	110: //Verifica se a reta indexada é a última criada
		IF NOT IHM.CutMode THEN
			IF PLC.CutLine = PLC.Grid THEN
				Auto.State := 118;
				ELSIF PLC.CutLine <> PLC.Grid THEN
					Auto.State := 111;
			END_IF
			ELSIF IHM.CutMode THEN
				IF PLC.CutLine = PLC.GridDesigner_LastLine THEN
					Auto.State := 118;
					ELSIF PLC.CutLine <> PLC.GridDesigner_LastLine THEN
						Auto.State := 111;
				END_IF
		END_IF
	
	111: //Passa para próxima reta
		PLC.CutLine := PLC.CutLine + 1;
		Auto.State := 30;
	
	118: //Recebe valor da última reta do eixo da altura ou primeira reta do eixo da largura
		IF NOT IHM.CutMode THEN
			PLC.CutLine := PLC.GridDesigner_LastLine;
			Auto.State := 119;
			ELSIF IHM.CutMode THEN
				PLC.CutLine := 21;
				Auto.State := 119;
		END_IF
	
	119: //Serra 90° ou 0° + Serra Ligada
		IF NOT IHM.CutMode THEN
			PLC.Axis[4].OperationDistance := 0;
			Auto.State := 120;
			ELSIF IHM.CutMode THEN
				PLC.Axis[4].OperationDistance := 90;
				Auto.State := 120;
		END_IF
	
	120: //Movimenta eixo W
		PLC.Axis[4].OperationStart := TRUE;
		IF NOT PLC.Axis[4].OperationDone THEN
			Auto.State := 121;
		END_IF
	
	121: //Aguarda movimentação do eixo
		IF PLC.Axis[4].OperationDone THEN
			PLC.Axis[4].OperationStart := FALSE;
			Auto.State := 122;
		END_IF
	
	122: //Posicão Zero Peça X (descontando borda de entrada) + Zero Peça Y da peça indexada
		IF NOT IHM.CutMode THEN
			PLC.Axis[1].OperationDistance := PLC.OrthogonalPieces[PLC.CutLine].LastVertexAbsX + (IHM.PrEntryEdgeX * -1);
			PLC.Axis[2].OperationDistance := PLC.OrthogonalPieces[PLC.CutLine].ZeroPieceY;
			PLC.Axis[1].OperationAbsolute := TRUE;
			PLC.Axis[2].OperationAbsolute := TRUE;
			Auto.State := 130;
			ELSIF IHM.CutMode THEN
				PLC.Axis[1].OperationDistance := PLC.OrthogonalPieces[PLC.CutLine].ZeroPieceX;
				PLC.Axis[2].OperationDistance := PLC.OrthogonalPieces[PLC.CutLine].ZeroPieceY + IHM.PrEntryEdgeY;
				PLC.Axis[1].OperationAbsolute := TRUE;
				PLC.Axis[2].OperationAbsolute := TRUE;
				Auto.State := 130;
		END_IF
	
	130: //Movimenta eixo X
		PLC.Axis[1].OperationStart := TRUE;
		IF NOT PLC.Axis[1].OperationDone THEN
			Auto.State := 131;
		END_IF
	
	131: //Movimenta eixo Y
		PLC.Axis[2].OperationStart := TRUE;
		IF NOT PLC.Axis[2].OperationDone THEN
			Auto.State := 132;
		END_IF
	
	132: //Aguarda movimento 90°/0° e movimentações de X e Y
		IF NOT IHM.CutMode AND PLC.Axis[4].Position = 0 OR IHM.CutMode AND PLC.Axis[4].Position = 90 THEN
			IF PLC.Axis[1].OperationDone AND PLC.Axis[2].OperationDone THEN
				PLC.Axis[1].OperationStart := FALSE;
				PLC.Axis[2].OperationStart := FALSE;
				Auto.State := 140;
			END_IF
		END_IF
	
	140: //Posição dentro da peça
		PLC.Axis[3].OperationDistance := IHM.PrInsidePiece;
		PLC.Axis[3].OperationAbsolute := TRUE;
		Auto.State := 150;
	
	150: //Movimenta eixo Z
		PLC.Axis[3].OperationStart := TRUE;
		IF NOT PLC.Axis[3].OperationDone THEN
			Auto.State := 151;
		END_IF
	
	151: //Aguarda movimentação do eixo
		IF PLC.Axis[3].OperationDone THEN
			PLC.Axis[3].OperationStart := FALSE;
			Auto.State := 160;
		END_IF
	
	160: //Deslocamento da largura (descontando bordas de entrada e saída) da peça indexada
		IF NOT IHM.CutMode THEN
			PLC.Axis[1].OperationDistance := (PLC.OrthogonalPieces[PLC.CutLine].Lenght * -1) + IHM.PrEntryEdgeX + IHM.PrLeadingEdgeX;
			PLC.Axis[1].OperationAbsolute := FALSE;
			Auto.State := 170;
			ELSIF IHM.CutMode THEN
				PLC.Axis[2].OperationDistance := PLC.OrthogonalPieces[PLC.CutLine].Lenght + (IHM.PrEntryEdgeY * -1) + (IHM.PrLeadingEdgeY * -1);
				PLC.Axis[2].OperationAbsolute := FALSE;
				Auto.State := 170;
		END_IF
	
	170: //Movimenta X ou Y
		IF NOT IHM.CutMode THEN
			PLC.Axis[1].OperationStart := TRUE;
			IF NOT PLC.Axis[1].OperationDone THEN
				Auto.State := 171;
			END_IF
			ELSIF IHM.CutMode THEN
				PLC.Axis[2].OperationStart := TRUE;
				IF NOT PLC.Axis[2].OperationDone THEN
					Auto.State := 171;
				END_IF
		END_IF
	
	171: //Aguarda movimentação X ou Y
		IF NOT IHM.CutMode AND PLC.Axis[1].OperationDone THEN
			PLC.Axis[1].OperationStart := FALSE;
			Auto.State := 180;
			ELSIF IHM.CutMode AND PLC.Axis[2].OperationDone THEN
				PLC.Axis[2].OperationStart := FALSE;
				Auto.State := 180;
		END_IF
	
	180: //Posição fora da peça
		PLC.Axis[3].OperationDistance := IHM.PrOutsidePiece;
		PLC.Axis[3].OperationAbsolute := TRUE;
		Auto.State := 190;
	
	190: //Movimenta eixo Z
		PLC.Axis[3].OperationStart := TRUE;
		IF NOT PLC.Axis[3].OperationDone THEN
			Auto.State := 191;
		END_IF
	
	191: //Aguarda movimentação do eixo
		IF PLC.Axis[3].OperationDone THEN
			PLC.Axis[3].OperationStart := FALSE;
			Auto.State := 200;
		END_IF
	
	200: //Verifica se a reta indexada é a primeira
		IF NOT IHM.CutMode THEN
			IF PLC.CutLine = 0 THEN
				Auto.State := 1000;
				ELSIF PLC.CutLine <> 0 THEN
					Auto.State := 201;
			END_IF
			ELSIF IHM.CutMode THEN
				IF PLC.CutLine = PLC.Grid THEN
					Auto.State := 1000;
					ELSIF PLC.CutLine <> PLC.Grid THEN
						Auto.State := 202;
				END_IF
		END_IF
	
	201: //Passa para reta anterior
		PLC.CutLine := PLC.CutLine - 1;
		Auto.State := 122;
	
	202: //Passa para reta peça
		PLC.CutLine := PLC.CutLine + 1;
		Auto.State := 122;
	
	999: //Abortar rotina
		Automatic_Abort();
	
	1000: //Finalizar rotina
		Automatic_Done();
END_CASE
                    
END_ACTION

ACTION Cutting_Corner:
                      (*Condição para habilitar modo automático*)
IF PLC.Machine = States.Manual THEN
	IF IHM.btStart OR PLC.IO.Start THEN
		Auto.Start := TRUE;
		PLC.Machine := States.Automatic;
		Auto.State := 1;
	END_IF
	(*Condição para parar processo*)
	ELSIF PLC.Machine = States.Automatic THEN
		IF IHM.btStop OR PLC.IO.Stop OR PLC.Axis[1].Error OR PLC.Axis[2].Error OR PLC.Axis[3].Error OR PLC.Axis[4].Error THEN
			Auto.State := 999;
		END_IF
END_IF

(*Rotina de corte corner [L]*)
CASE Auto.State OF
	1: //Estado rodando
		Automatic_Running();
	
	2: //Reseta variaveis
		AutomaticCorner_Reverse := FALSE;
		PLC.CutStraight := 0;
		AutomaticCorner_CuttingStep := 0;
		Auto.State := 10;
	
	10: //Posição fora da peça
		PLC.Axis[3].OperationDistance := IHM.PrOutsidePiece;
		PLC.IO.SawSpin := TRUE;
		PLC.Axis[3].OperationAbsolute := TRUE;
		Auto.State := 11;
	
	11: //Movimenta eixo Z
		PLC.Axis[3].OperationStart := TRUE;
		IF NOT PLC.Axis[3].OperationDone THEN
			Auto.State := 12;
		END_IF
	
	12: //Aguarda movimntação do eixo
		IF PLC.Axis[3].OperationDone THEN
			PLC.Axis[3].OperationStart := FALSE;
			Auto.State := 20;
		END_IF
	
	20: //Serra 90°
		PLC.Axis[4].OperationDistance := 90;
		Auto.State := 21;
	
	21: //Movimenta eixo W
		PLC.Axis[4].OperationStart := TRUE;
		IF NOT PLC.Axis[4].OperationDone THEN
			Auto.State := 22;
		END_IF
	
	22: //Aguarda movimentação do eixo
		IF PLC.Axis[4].OperationDone THEN
			PLC.Axis[4].OperationStart := FALSE;
			Auto.State := 30;
		END_IF
	
	30: //Posicão Zero Peça X + Zero Peça Y (descontando borda de entrada) da peça indexada
		IF NOT AutomaticCorner_HorizontalCutting THEN
			PLC.Axis[1].OperationDistance := PLC.CornerPieces[PLC.CutStraight].ZeroPieceX;
			PLC.Axis[2].OperationDistance := PLC.CornerPieces[PLC.CutStraight].ZeroPieceY + PLC.CornerPieces[PLC.CutStraight].EntryEdge;
			PLC.Axis[1].OperationAbsolute := TRUE;
			PLC.Axis[2].OperationAbsolute := TRUE;
			Auto.State := 40;
			ELSIF AutomaticCorner_HorizontalCutting THEN
				PLC.Axis[1].OperationDistance := PLC.CornerPieces[PLC.CutStraight].LastVertexAbsX + (PLC.CornerPieces[PLC.CutStraight].EntryEdge * -1);
				PLC.Axis[2].OperationDistance := PLC.CornerPieces[PLC.CutStraight].ZeroPieceY;
				PLC.Axis[1].OperationAbsolute := TRUE;
				PLC.Axis[2].OperationAbsolute := TRUE;
				Auto.State := 40;
		END_IF
	
	40: //Movimenta eixo X
		PLC.Axis[1].OperationStart := TRUE;
		IF NOT PLC.Axis[1].OperationDone THEN
			Auto.State := 41;
		END_IF
	
	41: //Movimenta eixo Y
		PLC.Axis[2].OperationStart := TRUE;
		IF NOT PLC.Axis[2].OperationDone THEN
			Auto.State := 42;
		END_IF
	
	42: //Aguardaserra 90° ou 0° e movimentações do eixo X e Y
		IF (NOT AutomaticCorner_HorizontalCutting AND PLC.Axis[4].Position = 90 AND PLC.Axis[1].OperationDone AND PLC.Axis[2].OperationDone) OR (AutomaticCorner_HorizontalCutting AND PLC.Axis[4].Position = 90 AND PLC.Axis[1].OperationDone AND PLC.Axis[2].OperationDone) THEN
			PLC.Axis[1].OperationStart := FALSE;
			PLC.Axis[2].OperationStart := FALSE;
			Auto.State := 50;
		END_IF
	
	50: //Posição dentro da peça
		PLC.Axis[3].OperationDistance := IHM.PrInsidePiece;
		PLC.Axis[3].OperationAbsolute := TRUE;
		Auto.State := 60;
	
	60: //Movimenta eixo Z
		PLC.Axis[3].OperationStart := TRUE;
		IF NOT PLC.Axis[3].OperationDone THEN
			Auto.State := 61;
		END_IF
	
	61: //Aguarda movimentação do eixo
		IF PLC.Axis[3].OperationDone THEN
			PLC.Axis[3].OperationStart := FALSE;
			Auto.State := 70;
		END_IF
	
	70: //Deslocamento da altura (descontando bordas de entrada e saída) da peça indexada
		IF NOT AutomaticCorner_HorizontalCutting THEN
			PLC.Axis[2].OperationDistance := PLC.CornerPieces[PLC.CutStraight].Height + (PLC.CornerPieces[PLC.CutStraight].EntryEdge * -1) + (PLC.CornerPieces[PLC.CutStraight].LeadingEdge * -1);
			PLC.Axis[2].OperationAbsolute := FALSE;
			Auto.State := 80;
			ELSIF AutomaticCorner_HorizontalCutting THEN
				PLC.Axis[1].OperationDistance := (PLC.CornerPieces[PLC.CutStraight].Width * -1) + PLC.CornerPieces[PLC.CutStraight].EntryEdge + PLC.CornerPieces[PLC.CutStraight].LeadingEdge;
				PLC.Axis[1].OperationAbsolute := FALSE;
				Auto.State := 80;
		END_IF
	
	80: //Movimenta eixo X ou Y
		IF NOT AutomaticCorner_HorizontalCutting THEN
			PLC.Axis[2].OperationStart := TRUE;
			IF NOT PLC.Axis[2].OperationDone THEN
				Auto.State := 81;
			END_IF
			ELSIF AutomaticCorner_HorizontalCutting THEN
				PLC.Axis[1].OperationStart := TRUE;
				IF NOT PLC.Axis[1].OperationDone THEN
					Auto.State := 81;
				END_IF
		END_IF
	
	81: //Aguarda movimentação X ou Y
		IF NOT AutomaticCorner_HorizontalCutting AND PLC.Axis[2].OperationDone THEN
			PLC.Axis[2].OperationStart := FALSE;
			Auto.State := 90;
			ELSIF AutomaticCorner_HorizontalCutting AND PLC.Axis[1].OperationDone THEN
				PLC.Axis[1].OperationStart := FALSE;
				Auto.State := 90;
		END_IF
	
	90: //Posição fora de peça
		PLC.Axis[3].OperationDistance := IHM.PrOutsidePiece;
		PLC.Axis[3].OperationAbsolute := TRUE;
		Auto.State := 100;
	
	100: //Movimenta eixo Z
		PLC.Axis[3].OperationStart := TRUE;
		IF NOT PLC.Axis[3].OperationDone THEN
			Auto.State := 101;
		END_IF
	
	101: //Aguarda movimentação do eixo
		IF PLC.Axis[3].OperationDone THEN
			PLC.Axis[3].OperationStart := FALSE;
			Auto.State := 110;
		END_IF
	
	110: //Verifica espelhamento
		IF NOT IHM.CreationCorner_MirrorCorner THEN
			IF NOT AutomaticCorner_HorizontalCutting AND PLC.CutStraight = 2 THEN
				Auto.State := 111;
			END_IF
			IF (NOT AutomaticCorner_HorizontalCutting AND PLC.CutStraight <> 2) OR (AutomaticCorner_HorizontalCutting AND PLC.CutStraight <> 5) THEN
				Auto.State := 120;
			END_IF
			IF AutomaticCorner_HorizontalCutting AND PLC.CutStraight = 5 THEN
				Auto.State := 1000;
			END_IF
			ELSIF IHM.CreationCorner_MirrorCorner THEN
				IF NOT AutomaticCorner_HorizontalCutting AND PLC.CutStraight = 3 THEN
					Auto.State := 111;
				END_IF
				IF (NOT AutomaticCorner_HorizontalCutting AND PLC.CutStraight <> 3) OR (AutomaticCorner_HorizontalCutting AND PLC.CutStraight <> 8) THEN
					Auto.State := 120;
				END_IF
				IF AutomaticCorner_HorizontalCutting AND PLC.CutStraight = 8 THEN
					Auto.State := 1000;
				END_IF
		END_IF
	
	111: //Passa para próxima reta e gira serra para 0°
		AutomaticCorner_HorizontalCutting := TRUE;
		PLC.Axis[4].OperationDistance := 0;
		Auto.State := 112;
	
	112: //Movimenta eixo W
		PLC.Axis[4].OperationStart := TRUE;
		IF NOT PLC.Axis[4].OperationDone THEN
			Auto.State := 113;
		END_IF
	
	113: //Aguarda movimentação do eixo
		IF PLC.Axis[4].OperationDone THEN
			PLC.Axis[4].OperationStart := FALSE;
			Auto.State := 120;
		END_IF
	
	120: //Passa para próxima reta
		PLC.CutStraight := PLC.CutStraight + 1;
		Auto.State := 30;
	
	999: //Abortar rotina
		Automatic_Abort();
	
	1000: //Finaliza rotina
		Automatic_Done();
END_CASE
                    
END_ACTION

ACTION Cutting_Forms:
                      (*Condição para habilitar modo automático*)
IF PLC.Machine = States.Manual THEN
	IF IHM.btStart OR PLC.IO.Start THEN
		Auto.Start := TRUE;
		PLC.Machine := States.Automatic;
		Auto.State := 1;
	END_IF
	(*Condição para parar processo*)
	ELSIF PLC.Machine = States.Automatic THEN
		IF IHM.btStop OR PLC.IO.Stop OR PLC.Axis[1].Error OR PLC.Axis[2].Error OR PLC.Axis[3].Error OR PLC.Axis[4].Error THEN
			Auto.State := 999;
		END_IF
END_IF

(*Rotina de corte Formas*)
CASE Auto.State OF
	1: //Estado rodando
		Automatic_Running();
	
	2: //Reseta variaveis
		AutomaticForms_Segaments := 0;
		Auto.State := 10;
	
	10: //Posição fora da peça
		PLC.Axis[3].OperationDistance := IHM.PrOutsidePiece;
		PLC.Axis[3].OperationAbsolute := TRUE;
		PLC.IO.SawSpin := TRUE;
		Auto.State := 11;
	
	11: //Movimenta eixo Z
		PLC.Axis[3].OperationStart := TRUE;
		IF NOT PLC.Axis[3].OperationDone THEN
			Auto.State := 12;
		END_IF
	
	12: //Aguarda movimentação do eixo
		IF PLC.Axis[3].OperationDone THEN
			PLC.Axis[3].OperationStart := FALSE;
			Auto.State := 20;
		END_IF
	
	20: //Verifica qual figura foi selecionada
		IF IHM.Figure = 1 THEN
			Auto.State := 30; //Quadrado/Retangulo
			ELSIF IHM.Figure = 2 THEN
				Auto.State := 70; //Circulo
				ELSIF IHM.Figure = 3 THEN
					Auto.State := 50; //Hexagono
					ELSIF IHM.Figure = 4 THEN
						Auto.State := 60; //Triangulo
		END_IF

(*-----------------QUADRADO-----------------*)	
	
	30: //Gira serra 90°
		PLC.Axis[4].OperationDistance := 90;
		Auto.State := 31;
		
	31: //Movimenta eixo W
		PLC.Axis[4].OperationStart := TRUE;
		IF NOT PLC.Axis[4].OperationDone THEN
			Auto.State := 32;
		END_IF
	
	32: //Aguarda movimentação do eixo
		IF PLC.Axis[4].OperationDone THEN
			PLC.Axis[4].OperationStart := FALSE;
			Auto.State := 33;
		END_IF
	
	33: //Posição zero peça
		IF AutomaticForms_Segaments = 0 THEN
			PLC.Axis[1].OperationDistance := PLC.FormsSquare.ZeroPieceX;
			PLC.Axis[2].OperationDistance := PLC.FormsSquare.ZeroPieceY + IHM.PrEntryEdgeY;
			PLC.Axis[1].OperationAbsolute := TRUE;
			PLC.Axis[2].OperationAbsolute := TRUE;
			Auto.State := 34;
			ELSIF AutomaticForms_Segaments = 1 THEN
				PLC.Axis[1].OperationDistance := PLC.FormsSquare.LastVertexAbsX + IHM.SawThickness;
				PLC.Axis[2].OperationDistance := PLC.FormsSquare.ZeroPieceY + IHM.PrEntryEdgeY;
				PLC.Axis[1].OperationAbsolute := TRUE;
				PLC.Axis[2].OperationAbsolute := TRUE;
				Auto.State := 34;
		END_IF
	
	34: //Movimenta eixo X
		PLC.Axis[1].OperationStart := TRUE;
		IF NOT PLC.Axis[1].OperationDone THEN
			Auto.State := 35;
		END_IF
	
	35: //Movimenta eixo Y
		PLC.Axis[2].OperationStart := TRUE;
		IF NOT PLC.Axis[2].OperationDone THEN
			Auto.State := 36;
		END_IF
	
	36: //Aguarda movimento dos eixos e posição da serra 90°
		IF PLC.Axis[1].OperationDone AND PLC.Axis[2].OperationDone AND PLC.Axis[4].Position = 90 THEN
			PLC.Axis[1].OperationStart := FALSE;
			PLC.Axis[2].OperationStart := FALSE;
			Auto.State := 37;
		END_IF
	
	37: //Posição dentro da peça
		PLC.Axis[3].OperationDistance := IHM.PrInsidePiece;
		PLC.Axis[3].OperationAbsolute := TRUE;
		Auto.State := 38;
	
	38: //Movimenta eixo Z
		PLC.Axis[3].OperationStart := TRUE;
		IF NOT PLC.Axis[3].OperationDone THEN
			Auto.State := 39;
		END_IF
	
	39: //Aguarda movimentação do eixo
		IF PLC.Axis[3].OperationDone THEN
			PLC.Axis[3].OperationStart := FALSE;
			Auto.State := 40;
		END_IF
	
	40: //Deslocamento da altura
		PLC.Axis[2].OperationDistance := PLC.FormsSquare.Height + (IHM.PrEntryEdgeY * -1) + (IHM.PrLeadingEdgeY * -1);
		Auto.State := 41;
	
	41: //Movimenta eixo Y
		PLC.Axis[2].OperationStart := TRUE;
		IF NOT PLC.Axis[2].OperationDone THEN
			Auto.State := 42;
		END_IF
	
	42: //Aguarda movimento do eixo
		IF PLC.Axis[2].OperationDone THEN
			PLC.Axis[2].OperationStart := FALSE;
			Auto.State := 43;
		END_IF
	
	43: //Posição fora da peça
		PLC.Axis[3].OperationDistance := IHM.PrOutsidePiece;
		PLC.Axis[3].OperationAbsolute := TRUE;
		Auto.State := 44;
	
	44: //Movimento eixo Z
		PLC.Axis[3].OperationStart := TRUE;
		IF NOT PLC.Axis[3].OperationDone THEN
			Auto.State := 45;
		END_IF
	
	45: //Aguarda movimento do eixo
		IF PLC.Axis[3].OperationDone THEN
			PLC.Axis[3].OperationStart := FALSE;
			Auto.State := 46;
		END_IF
	
	46: //Soma na indexadora
		AutomaticForms_Segaments := AutomaticForms_Segaments + 1;
		Auto.State := 47;
	
	47: //Verifica se é o primeiro ou segundo corte
		IF AutomaticForms_Segaments = 2 THEN
			Auto.State := 48;
			ELSIF AutomaticForms_Segaments = 1 THEN
				Auto.State := 33;
		END_IF
	
	48: //Gira serra 0°
		PLC.Axis[4].OperationDistance := 0;
		Auto.State := 49;
		
	49: //Movimenta eixo W
		PLC.Axis[4].OperationStart := TRUE;
		IF NOT PLC.Axis[4].OperationDone THEN
			Auto.State := 50;
		END_IF
	
	50: //Aguarda movimentação do eixo
		IF PLC.Axis[4].OperationDone THEN
			PLC.Axis[4].OperationStart := FALSE;
			Auto.State := 51;
		END_IF
	
	51: //Posição zero peça
		IF AutomaticForms_Segaments = 2 THEN
			PLC.Axis[1].OperationDistance := PLC.FormsSquare.ZeroPieceX + IHM.PrEntryEdgeX;
			PLC.Axis[2].OperationDistance := PLC.FormsSquare.ZeroPieceY;
			Auto.State := 52;
			ELSIF AutomaticForms_Segaments = 3 THEN
				PLC.Axis[1].OperationDistance := PLC.FormsSquare.ZeroPieceX + IHM.PrEntryEdgeX;
				PLC.Axis[2].OperationDistance := PLC.FormsSquare.LastVertexAbsY + IHM.SawThickness;
				PLC.Axis[1].OperationAbsolute := TRUE;
				PLC.Axis[2].OperationAbsolute := TRUE;
				Auto.State := 52;
		END_IF
	
	52: //Movimenta eixo X
		PLC.Axis[1].OperationStart := TRUE;
		IF NOT PLC.Axis[1].OperationDone THEN
			Auto.State := 53;
		END_IF
	
	53: //Movimenta eixo Y
		PLC.Axis[2].OperationStart := TRUE;
		IF NOT PLC.Axis[2].OperationDone THEN
			Auto.State := 54;
		END_IF
	
	54: //Aguarda movimento dos eixos e posição da serra 0°
		IF PLC.Axis[1].OperationDone AND PLC.Axis[2].OperationDone AND PLC.Axis[4].Position = 0 THEN
			PLC.Axis[1].OperationStart := FALSE;
			PLC.Axis[2].OperationStart := FALSE;
			Auto.State := 55;
		END_IF
	
	55: //Posição dentro da peça
		PLC.Axis[3].OperationDistance := IHM.PrInsidePiece;
		PLC.Axis[3].OperationAbsolute := TRUE;
		Auto.State := 56;
	
	56: //Movimenta eixo Z
		PLC.Axis[3].OperationStart := TRUE;
		IF NOT PLC.Axis[3].OperationDone THEN
			Auto.State := 57;
		END_IF
	
	57: //Aguarda movimentação do eixo
		IF PLC.Axis[3].OperationDone THEN
			PLC.Axis[3].OperationStart := FALSE;
			Auto.State := 58;
		END_IF
	
	58: //Deslocamento da largura
		PLC.Axis[1].OperationDistance := PLC.FormsSquare.Width + (IHM.PrEntryEdgeX * -1) + (IHM.PrLeadingEdgeX * -1);
		Auto.State := 59;
	
	59: //Movimenta eixo Y
		PLC.Axis[1].OperationStart := TRUE;
		IF NOT PLC.Axis[1].OperationDone THEN
			Auto.State := 60;
		END_IF
	
	60: //Aguarda movimento do eixo
		IF PLC.Axis[1].OperationDone THEN
			PLC.Axis[1].OperationStart := FALSE;
			Auto.State := 61;
		END_IF
	
	61: //Posição fora da peça
		PLC.Axis[3].OperationDistance := IHM.PrOutsidePiece;
		PLC.Axis[3].OperationAbsolute := TRUE;
		Auto.State := 62;
	
	62: //Movimento eixo Z
		PLC.Axis[3].OperationStart := TRUE;
		IF NOT PLC.Axis[3].OperationDone THEN
			Auto.State := 63;
		END_IF
	
	63: //Aguarda movimento do eixo
		IF PLC.Axis[3].OperationDone THEN
			PLC.Axis[3].OperationStart := FALSE;
			Auto.State := 64;
		END_IF
	
	64: //Soma no indexador
		AutomaticForms_Segaments := AutomaticForms_Segaments + 1;
		Auto.State := 65;
	
	65: //Verifica se é o primeiro ou segundo corte
		IF AutomaticForms_Segaments = 4 THEN
			Auto.State := 1000;
			ELSIF AutomaticForms_Segaments = 3 THEN
				Auto.State := 51;
		END_IF
	
(*-----------------CIRCULO-----------------*)		
	
	70: //Gira serra 90°
		PLC.Axis[4].OperationDistance := 90;
		Auto.State := 71;
		
	71: //Movimenta eixo W
		PLC.Axis[4].OperationStart := TRUE;
		IF NOT PLC.Axis[4].OperationDone THEN
			Auto.State := 72;
		END_IF
	
	72: //Aguarda movimentação do eixo
		IF PLC.Axis[4].OperationDone THEN
			PLC.Axis[4].OperationStart := FALSE;
			Auto.State := 73;
		END_IF
	
	73: //Posição zero peça
		PLC.Axis[1].OperationDistance := PLC.FormsCircle.ZeroPieceX;
		PLC.Axis[2].OperationDistance := PLC.FormsCircle.Height / 2;
		PLC.Axis[1].OperationAbsolute := TRUE;
		PLC.Axis[2].OperationAbsolute := TRUE;
		Auto.State := 74;

	74: //Movimenta eixo X
		PLC.Axis[1].OperationStart := TRUE;
		IF NOT PLC.Axis[1].OperationDone THEN
			Auto.State := 75;
		END_IF
	
	75: //Movimenta eixo Y
		PLC.Axis[2].OperationStart := TRUE;
		IF NOT PLC.Axis[2].OperationDone THEN
			Auto.State := 76;
		END_IF
	
	76: //Aguarda movimento dos eixos e posição da serra 90°
		IF PLC.Axis[1].OperationDone AND PLC.Axis[2].OperationDone AND PLC.Axis[4].Position = 90 THEN
			PLC.Axis[1].OperationStart := FALSE;
			PLC.Axis[2].OperationStart := FALSE;
			Auto.State := 77;
		END_IF
	
	77: //Posição dentro da peça
		PLC.Axis[3].OperationDistance := IHM.PrInsidePiece;
		PLC.Axis[3].OperationAbsolute := TRUE;
		Auto.State := 78;
	
	78: //Movimenta eixo Z
		PLC.Axis[3].OperationStart := TRUE;
		IF NOT PLC.Axis[3].OperationDone THEN
			Auto.State := 79;
		END_IF
	
	79: //Aguarda movimentação do eixo
		IF PLC.Axis[3].OperationDone THEN
			PLC.Axis[3].OperationStart := FALSE;
			Auto.State := 80;
		END_IF
	
	80: //Primeira posição
		PLC.OperationAuxPos[0] := PLC.FormsCircle.Width / 2;
		PLC.OperationAuxPos[1] := PLC.FormsCircle.Height / 2;
		PLC.OperationEndPos[0] := PLC.FormsCircle.Width / 2;
		PLC.OperationEndPos[1] := PLC.FormsCircle.Height;
		Auto.State := 81;
	
	81: //Movimenta eixo X e Y
		PLC.OperationCirleStart := TRUE;
		IF NOT PLC.OperationCircleDone THEN
			Auto.State := 82;
		END_IF
	
	82: //Aguarda movimento
		IF PLC.OperationCircleDone THEN
			PLC.OperationCirleStart := FALSE;
			Auto.State := 83;
		END_IF
	
	83: //Segunda posição
		PLC.OperationAuxPos[0] := PLC.FormsCircle.Width / 2;
		PLC.OperationAuxPos[1] := PLC.FormsCircle.Height / 2;
		PLC.OperationEndPos[0] := PLC.FormsCircle.Width;
		PLC.OperationEndPos[1] := PLC.FormsCircle.Height / 2;
		Auto.State := 84;
	
	84: //Movimenta eixo X e Y
		PLC.OperationCirleStart := TRUE;
		IF NOT PLC.OperationCircleDone THEN
			Auto.State := 85;
		END_IF
	
	85: //Aguarda movimento
		IF PLC.OperationCircleDone THEN
			PLC.OperationCirleStart := FALSE;
			Auto.State := 86;
		END_IF
	
	86: //Terceira posição
		PLC.OperationAuxPos[0] := PLC.FormsCircle.Width / 2;
		PLC.OperationAuxPos[1] := PLC.FormsCircle.Height / 2;
		PLC.OperationEndPos[0] := PLC.FormsCircle.Width / 2;
		PLC.OperationEndPos[1] := PLC.FormsCircle.ZeroPieceY;
		Auto.State := 87;
	
	87: //Movimenta eixo X e Y
		PLC.OperationCirleStart := TRUE;
		IF NOT PLC.OperationCircleDone THEN
			Auto.State := 88;
		END_IF
	
	88: //Aguarda movimento
		IF PLC.OperationCircleDone THEN
			PLC.OperationCirleStart := FALSE;
			Auto.State := 89;
		END_IF
	
	89: //Quarta posição
		PLC.OperationAuxPos[0] := PLC.FormsCircle.Width / 2;
		PLC.OperationAuxPos[1] := PLC.FormsCircle.Height / 2;
		PLC.OperationEndPos[0] := PLC.FormsCircle.ZeroPieceX;
		PLC.OperationEndPos[1] := PLC.FormsCircle.Height / 2;
		Auto.State := 90;
	
	90: //Movimenta eixo X e Y
		PLC.OperationCirleStart := TRUE;
		IF NOT PLC.OperationCircleDone THEN
			Auto.State := 91;
		END_IF
	
	91: //Aguarda movimento
		IF PLC.OperationCircleDone THEN
			PLC.OperationCirleStart := FALSE;
			Auto.State := 92;
		END_IF
	
	92: //Posição fora da peça
		PLC.Axis[3].OperationDistance := IHM.PrOutsidePiece;
		PLC.Axis[3].OperationAbsolute := TRUE;
		Auto.State := 93;
	
	93: //Movimenta eixo Z
		PLC.Axis[3].OperationStart := TRUE;
		IF NOT PLC.Axis[3].OperationDone THEN
			Auto.State := 94;
		END_IF
	
	94: //Aguarda movimentação do eixo
		IF PLC.Axis[3].OperationDone THEN
			PLC.Axis[3].OperationStart := FALSE;
			Auto.State := 1000;
		END_IF
	
(*-----------------HEXAGONO-----------------*)	
	
	100:
		;

	999: //Abortar rotina
		Automatic_Abort();
END_CASE
                    
END_ACTION

METHOD SetPoint
  VAR_INPUT
    Execute : BOOL;
  END_VAR
                        (*Define novo ponto zero*)
FB_Setpoint[1](Axis := Axis1, Execute := Execute, Position := 0);
FB_Setpoint[2](Axis := Axis2, Execute := Execute, Position := 0);
FB_Setpoint[3](Axis := Axis3, Execute := Execute, Position := 0);
                      
END_METHOD

METHOD GoToZero
  VAR_INPUT
    Execute : BOOL;
  END_VAR
                        (*Condição para retornar para zero*)
IF Execute THEN
	//Posição para os eixos
	PLC.Axis[1].OperationDistance := 0;
	PLC.Axis[2].OperationDistance := 0;
	PLC.Axis[3].OperationDistance := 0;
	//Executa eixos
	PLC.Axis[1].OperationStart := TRUE;
	PLC.Axis[2].OperationStart := TRUE;
	PLC.Axis[3].OperationStart := TRUE;
	//Modo Absoluto
	PLC.Axis[1].OperationAbsolute := TRUE;
	PLC.Axis[2].OperationAbsolute := TRUE;
	PLC.Axis[3].OperationAbsolute := TRUE;
	(*Condição para finalizar retorno*)
	IF PLC.Axis[1].OperationDone AND PLC.Axis[2].OperationDone AND PLC.Axis[3].OperationDone THEN
		//Desabilita execução dos eixos
		PLC.Axis[1].OperationStart := FALSE;
		PLC.Axis[2].OperationStart := FALSE;
		PLC.Axis[3].OperationStart := FALSE;
		PLC.Axis[1].OperationAbsolute := FALSE;
		PLC.Axis[2].OperationAbsolute := FALSE;
		PLC.Axis[3].OperationAbsolute := FALSE;
		//Desabilita condição para retorno
		IHM.btGoToZero := FALSE;
	END_IF
	(*Condição para parar retorno*)
	IF IHM.btStop OR PLC.IO.Stop THEN
		//Desabilita execução dos eixos
		PLC.Axis[1].OperationStart := FALSE;
		PLC.Axis[2].OperationStart := FALSE;
		PLC.Axis[3].OperationStart := FALSE;
		PLC.Axis[1].OperationAbsolute := FALSE;
		PLC.Axis[2].OperationAbsolute := FALSE;
		PLC.Axis[3].OperationAbsolute := FALSE;
		//Desabilita condição para retorno
		IHM.btGoToZero := FALSE;
	END_IF
END_IF
                      
END_METHOD

METHOD RotateSaw
  VAR_INPUT
    Execute : BOOL;
  END_VAR
                        (*Condição para girar a serra*)
IF Execute THEN
	//Posição para o eixo
	PLC.Axis[4].OperationDistance := IHM.RotateValue;
	//Executa eixos
	PLC.Axis[4].OperationStart := TRUE;
	(*Condição para finalizar função*)
	IF PLC.Axis[4].OperationDone THEN
		//Desabilita execução dos eixos
		PLC.Axis[4].OperationStart := FALSE;
		//Desabilita condição para retorno
		IHM.btRotateSaw := FALSE;
	END_IF
	(*Condição para parar retorno*)
	IF IHM.btStop OR PLC.IO.Stop THEN
		//Desabilita execução dos eixos
		PLC.Axis[4].OperationStart := FALSE;
		//Desabilita condição para retorno
		IHM.btRotateSaw := FALSE;
	END_IF
END_IF
                      
END_METHOD

METHOD TableUp
  VAR_INPUT
    Execute : BOOL;
  END_VAR
                        IF Execute AND PLC.IO.SsMesaBaixa THEN
	PLC.IO.SobeMesa := TRUE;
	ELSE
		PLC.IO.SobeMesa := FALSE;
END_IF
                      
END_METHOD

METHOD Input
  VAR_INPUT
    dwInput : DWORD;
  END_VAR
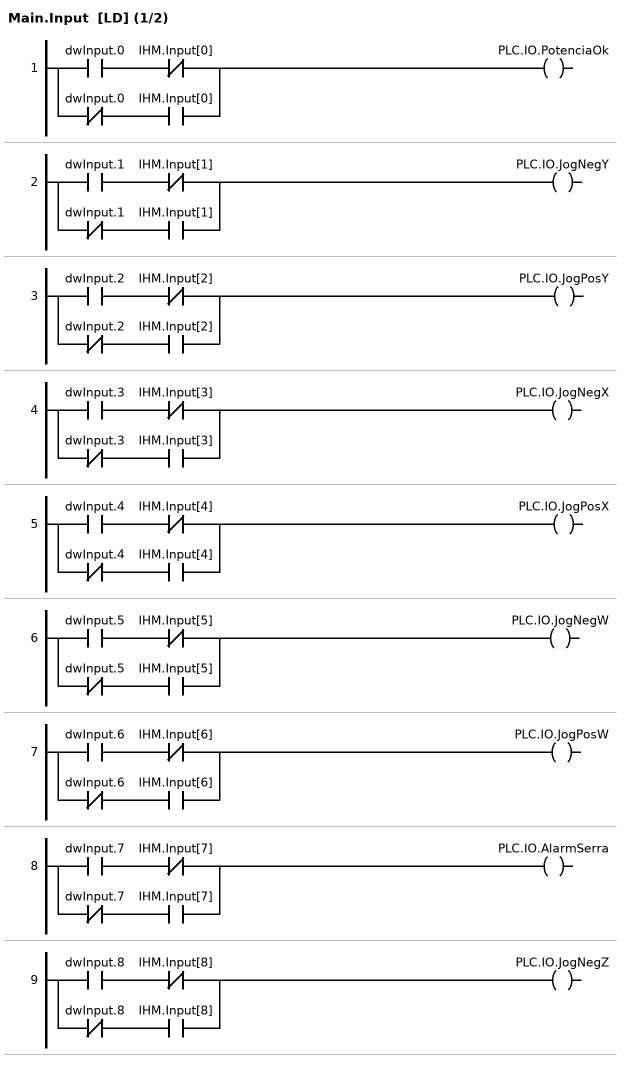
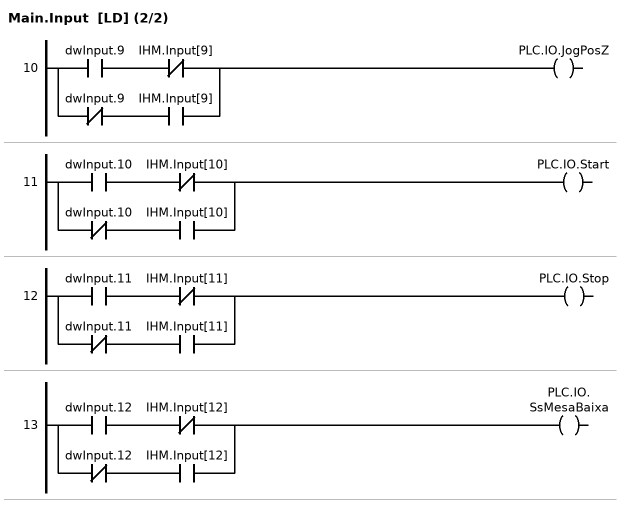
(* LD diagram, written out as Structured Text *)
(* Entrada 0 - Potencia OK *)

PLC.IO.PotenciaOk := dwInput.0 AND NOT IHM.Input[0] OR NOT dwInput.0 AND IHM.Input[0];
(* Entrada 1 - Movimento Negativo em Y *)

PLC.IO.JogNegY := dwInput.1 AND NOT IHM.Input[1] OR NOT dwInput.1 AND IHM.Input[1];
(* Entrada 2 - Movimento Positivo em Y *)

PLC.IO.JogPosY := dwInput.2 AND NOT IHM.Input[2] OR NOT dwInput.2 AND IHM.Input[2];
(* Entrada 3 - Movimento Negativo em X *)

PLC.IO.JogNegX := dwInput.3 AND NOT IHM.Input[3] OR NOT dwInput.3 AND IHM.Input[3];
(* Entrada 4 - Movimento Positivo em X *)

PLC.IO.JogPosX := dwInput.4 AND NOT IHM.Input[4] OR NOT dwInput.4 AND IHM.Input[4];
(* Entrada 5 - Movimento Negativo em W *)

PLC.IO.JogNegW := dwInput.5 AND NOT IHM.Input[5] OR NOT dwInput.5 AND IHM.Input[5];
(* Entrada 6 - Movimento Positivo em W *)

PLC.IO.JogPosW := dwInput.6 AND NOT IHM.Input[6] OR NOT dwInput.6 AND IHM.Input[6];
(* Entrada 7 - Alarme Serra *)

PLC.IO.AlarmSerra := dwInput.7 AND NOT IHM.Input[7] OR NOT dwInput.7 AND IHM.Input[7];
(* Entrada 8 - Movimento Negativo em Z *)

PLC.IO.JogNegZ := dwInput.8 AND NOT IHM.Input[8] OR NOT dwInput.8 AND IHM.Input[8];
(* Entrada 9 - Movimento Positivo em Z *)

PLC.IO.JogPosZ := dwInput.9 AND NOT IHM.Input[9] OR NOT dwInput.9 AND IHM.Input[9];
(* Entrada 10 - Botão Start *)

PLC.IO.Start := dwInput.10 AND NOT IHM.Input[10] OR NOT dwInput.10 AND IHM.Input[10];
(* Entrada 11 - Botão Stop *)

PLC.IO.Stop := dwInput.11 AND NOT IHM.Input[11] OR NOT dwInput.11 AND IHM.Input[11];
(* Entrada 12 - Sensor Mesa Baixa *)

PLC.IO.SsMesaBaixa := dwInput.12 AND NOT IHM.Input[12] OR NOT dwInput.12 AND IHM.Input[12];
END_METHOD

METHOD Output
  VAR_OUTPUT
    dwOutput : DWORD;
  END_VAR
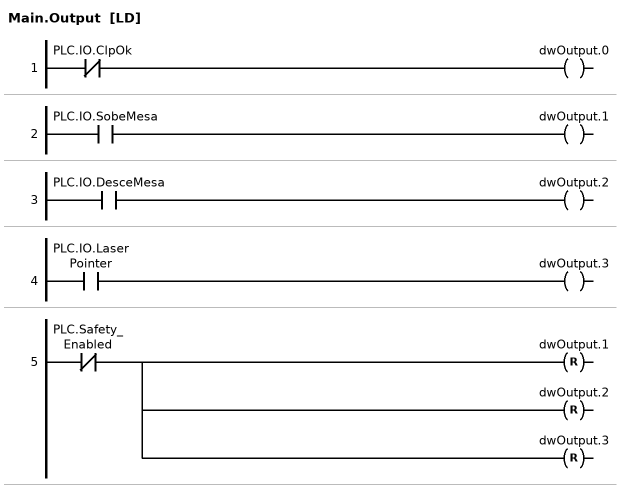
(* LD diagram, written out as Structured Text *)
(* Saida 0 - CLP Ok *)

dwOutput.0 := NOT PLC.IO.ClpOk;
(* Saida 1 - Sobe Mesa *)

dwOutput.1 := PLC.IO.SobeMesa;
(* Saida 2 - Desce Mesa *)

dwOutput.2 := PLC.IO.DesceMesa;
(* Saida 2 - Liga Laser Pointer *)

dwOutput.3 := PLC.IO.LaserPointer;
(* Reseta Saídas em caso de emergência *)

IF NOT PLC.Safety_Enabled THEN dwOutput.1 := FALSE; END_IF;
IF NOT PLC.Safety_Enabled THEN dwOutput.2 := FALSE; END_IF;
IF NOT PLC.Safety_Enabled THEN dwOutput.3 := FALSE; END_IF;
END_METHOD

METHOD TableDown
  VAR_INPUT
    Execute : BOOL;
  END_VAR
                        IF Execute AND NOT PLC.IO.SsMesaBaixa THEN
	PLC.IO.DesceMesa := TRUE;
	ELSE
		PLC.IO.DesceMesa := FALSE;
END_IF
                      
END_METHOD
END_PROGRAM

PROGRAM Motion
  VAR
    FB_Power : ARRAY[1..4] OF MC_Power;
    FB_Reset : ARRAY[1..4] OF MC_Reset;
    FB_Error : ARRAY[1..4] OF MC_ReadAxisError;
    FB_Jog : ARRAY[1..4] OF MC_Jog;
    FB_Absolute : ARRAY[1..4] OF MC_MoveAbsolute;
    FB_Relative : ARRAY[1..3] OF MC_MoveRelative;
    FB_Stop : ARRAY[1..4] OF MC_Stop;
    FB_Position : ARRAY[1..4] OF MC_ReadActualPosition;
    FB_Circular : LS_2AxisCircle;
  END_VAR

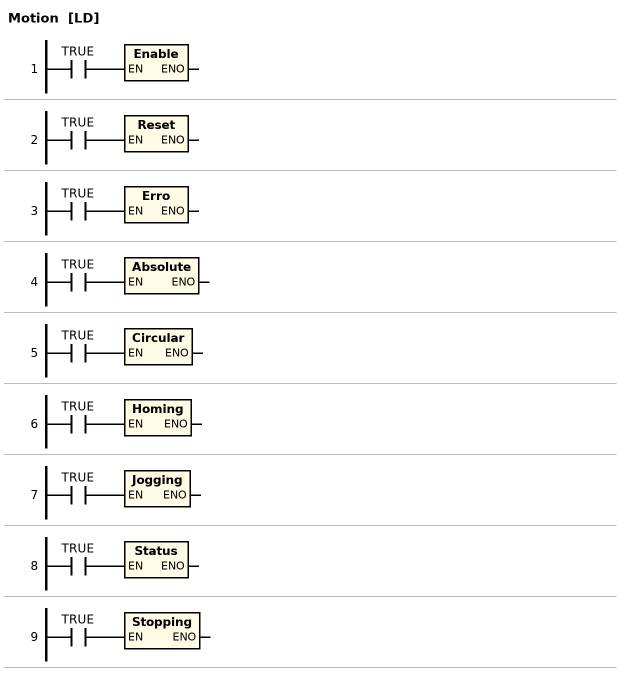
(* LD diagram, written out as Structured Text *)
(* Controle para habilitar os eixos *)

IF TRUE THEN Enable(); END_IF;
(* Controle para resetar os eixos *)

IF TRUE THEN Reset(); END_IF;
(* Controle de erros nos eixos *)

IF TRUE THEN Erro(); END_IF;
(* Controle de movimento absoluto dos eixos *)

IF TRUE THEN Absolute(); END_IF;

IF TRUE THEN Circular(); END_IF;
(* Controle de referência dos eixos *)

IF TRUE THEN Homing(); END_IF;
(* Controle de JOG dos eixos *)

IF TRUE THEN Jogging(); END_IF;
(* Status dos eixos *)

IF TRUE THEN Status(); END_IF;
(* Parada dos eixos *)

IF TRUE THEN Stopping(); END_IF;

ACTION Erro:
                      (*Informa erro nos eixos*)
FB_Error[1](Axis := Axis1, Enable := TRUE, AxisError => PLC.Axis[1].Error, AxisErrorID => PLC.Axis[1].ErrorID);
FB_Error[2](Axis := Axis2, Enable := TRUE, AxisError => PLC.Axis[2].Error, AxisErrorID => PLC.Axis[2].ErrorID);
FB_Error[3](Axis := Axis3, Enable := TRUE, AxisError => PLC.Axis[3].Error, AxisErrorID => PLC.Axis[3].ErrorID);
FB_Error[4](Axis := Axis4, Enable := TRUE, AxisError => PLC.Axis[4].Error, AxisErrorID => PLC.Axis[4].ErrorID);
                    
END_ACTION

ACTION Reset:
                      (*Reseta eixos*)
FB_Reset[1](Axis := Axis1, Execute := IHM.btReset AND PLC.Axis[1].Error);
FB_Reset[2](Axis := Axis2, Execute := IHM.btReset AND PLC.Axis[2].Error);
FB_Reset[3](Axis := Axis3, Execute := IHM.btReset AND PLC.Axis[3].Error);
FB_Reset[4](Axis := Axis4, Execute := IHM.btReset AND PLC.Axis[4].Error);
                    
END_ACTION

ACTION Enable:
                      (*Habilita eixos*)
FB_Power[1](Axis := Axis1, Enable := TRUE, bRegulatorOn := PLC.Safety_Enabled, bDriveStart := PLC.Safety_Enabled);
FB_Power[2](Axis := Axis2, Enable := TRUE, bRegulatorOn := PLC.Safety_Enabled, bDriveStart := PLC.Safety_Enabled);
FB_Power[3](Axis := Axis3, Enable := TRUE, bRegulatorOn := PLC.Safety_Enabled, bDriveStart := PLC.Safety_Enabled);
FB_Power[4](Axis := Axis4, Enable := TRUE, bRegulatorOn := PLC.Safety_Enabled, bDriveStart := PLC.Safety_Enabled);
                    
END_ACTION

ACTION Absolute:
                      (*Movimento absoluto para os eixos*)
FB_Absolute[1](	//Eixo 1
	Axis := Axis1,
	Execute := PLC.Axis[1].OperationStart,
	Position := PLC.Axis[1].OperationDistance,
	Velocity := PLC.Axis[1].OperationSpeed,
	Acceleration := PLC.Axis[1].Acceleration,
	Deceleration := PLC.Axis[1].Deceleration,
	Done => PLC.Axis[1].OperationDone);
	
FB_Absolute[2](	//Eixo 2
	Axis := Axis2,
	Execute := PLC.Axis[2].OperationStart,
	Position := PLC.Axis[2].OperationDistance,
	Velocity := PLC.Axis[2].OperationSpeed,
	Acceleration := PLC.Axis[2].Acceleration,
	Deceleration := PLC.Axis[2].Deceleration,
	Done => PLC.Axis[2].OperationDone);

FB_Absolute[3](	//Eixo 3
	Axis := Axis3,
	Execute := PLC.Axis[3].OperationStart,
	Position := PLC.Axis[3].OperationDistance,
	Velocity := PLC.Axis[3].OperationSpeed,
	Acceleration := PLC.Axis[3].Acceleration,
	Deceleration := PLC.Axis[3].Deceleration,
	Done => PLC.Axis[3].OperationDone);

FB_Absolute[4](	//Eixo 4
	Axis := Axis4,
	Execute := PLC.Axis[4].OperationStart,
	Position := PLC.Axis[4].OperationDistance,
	Velocity := PLC.Axis[4].OperationSpeed,
	Acceleration := PLC.Axis[4].Acceleration,
	Deceleration := PLC.Axis[4].Deceleration,
	Done => PLC.Axis[4].OperationDone);
                    
END_ACTION

ACTION Homing:
                      (*Homing dos eixos*)
PLC.FB_Homing[1](	//Eixo 1
	Axis := Axis1,
	fVelocitySlow := PLC.Axis[1].CreepSpeed,
	fVelocityFast := PLC.Axis[1].HomeSpeed,
	fAcceleration := PLC.Axis[1].Acceleration,
	fDeceleration := PLC.Axis[1].Deceleration,
	nDirection := PLC.Axis[1].HomeDirection,
	bReferenceSwitch := ,
	nHomingMode := SMC_HOMING_MODE.FAST_BSLOW_STOP_S,
	bDone => PLC.Axis[1].HomeDone);

PLC.FB_Homing[2](	//Eixo 2
	Axis := Axis2,
	fVelocitySlow := PLC.Axis[2].CreepSpeed,
	fVelocityFast := PLC.Axis[2].HomeSpeed,
	fAcceleration := PLC.Axis[2].Acceleration,
	fDeceleration := PLC.Axis[2].Deceleration,
	nDirection := PLC.Axis[2].HomeDirection,
	bReferenceSwitch := ,
	nHomingMode := SMC_HOMING_MODE.FAST_BSLOW_STOP_S,
	bDone => PLC.Axis[2].HomeDone);

PLC.FB_Homing[3](	//Eixo 3
	Axis := Axis3,
	fVelocitySlow := PLC.Axis[3].CreepSpeed,
	fVelocityFast := PLC.Axis[3].HomeSpeed,
	fAcceleration := PLC.Axis[3].Acceleration,
	fDeceleration := PLC.Axis[3].Deceleration,
	nDirection := PLC.Axis[3].HomeDirection,
	bReferenceSwitch := ,
	nHomingMode := SMC_HOMING_MODE.FAST_BSLOW_STOP_S,
	bDone => PLC.Axis[3].HomeDone);

PLC.FB_Homing[4](	//Eixo 4
	Axis := Axis4,
	fVelocitySlow := PLC.Axis[4].CreepSpeed,
	fVelocityFast := PLC.Axis[4].HomeSpeed,
	fAcceleration := PLC.Axis[4].Acceleration,
	fDeceleration := PLC.Axis[4].Deceleration,
	nDirection := PLC.Axis[4].HomeDirection,
	bReferenceSwitch := ,
	nHomingMode := SMC_HOMING_MODE.FAST_BSLOW_STOP_S,
	bDone => PLC.Axis[4].HomeDone);
                    
END_ACTION

ACTION Jogging:
                      (*JOG dos eixos*)
FB_Jog[1](	//Eixo 1
	Axis := Axis1,
	JogForward := PLC.Axis[1].JogFwd,
	JogBackward := PLC.Axis[1].JogRev,
	Velocity := PLC.Axis[1].ManualSpeed,
	Acceleration := PLC.Axis[1].Acceleration,
	Deceleration := PLC.Axis[1].Deceleration);

FB_Jog[2](	//Eixo 2
	Axis := Axis2,
	JogForward := PLC.Axis[2].JogFwd,
	JogBackward := PLC.Axis[2].JogRev,
	Velocity := PLC.Axis[2].ManualSpeed,
	Acceleration := PLC.Axis[2].Acceleration,
	Deceleration := PLC.Axis[2].Deceleration);

FB_Jog[3](	//Eixo 3
	Axis := Axis3,
	JogForward := PLC.Axis[3].JogFwd,
	JogBackward := PLC.Axis[3].JogRev,
	Velocity := PLC.Axis[3].ManualSpeed,
	Acceleration := PLC.Axis[3].Acceleration,
	Deceleration := PLC.Axis[3].Deceleration);

FB_Jog[4](	//Eixo 4
	Axis := Axis4,
	JogForward := PLC.Axis[4].JogFwd,
	JogBackward := PLC.Axis[4].JogRev,
	Velocity := PLC.Axis[4].ManualSpeed,
	Acceleration := PLC.Axis[4].Acceleration,
	Deceleration := PLC.Axis[4].Deceleration);

                    
END_ACTION

ACTION Status:
                      (*Posição dos eixos*)
FB_Position[1](	//Eixo 1
	Axis := Axis1,
	Enable := TRUE,
	Position => PLC.Axis[1].Position);

FB_Position[2](	//Eixo 2
	Axis := Axis2,
	Enable := TRUE,
	Position => PLC.Axis[2].Position);

FB_Position[3](	//Eixo 3
	Axis := Axis3,
	Enable := TRUE,
	Position => PLC.Axis[3].Position);

FB_Position[4](	//Eixo 4
	Axis := Axis4,
	Enable := TRUE,
	Position => PLC.Axis[4].Position);

                    
END_ACTION

ACTION Stopping:
                      (*Stop dos eixos*)
FB_Stop[1](	//Eixo 1
	Axis := Axis1,
	Execute := PLC.Axis[1].Stop OR PLC.IO.Stop,
	Deceleration := PLC.Axis[1].Deceleration);

FB_Stop[2](	//Eixo 2
	Axis := Axis2,
	Execute := PLC.Axis[2].Stop OR PLC.IO.Stop,
	Deceleration := PLC.Axis[2].Deceleration);

FB_Stop[3](	//Eixo 3
	Axis := Axis3,
	Execute := PLC.Axis[3].Stop OR PLC.IO.Stop,
	Deceleration := PLC.Axis[3].Deceleration);

FB_Stop[4](	//Eixo 4
	Axis := Axis4,
	Execute := PLC.Axis[4].Stop OR PLC.IO.Stop,
	Deceleration := PLC.Axis[4].Deceleration);
                    
END_ACTION

ACTION Relative:
                      (*Movimento absoluto para os eixos*)
FB_Relative[1]( //Eixo 1
	Axis := Axis1,
	Execute := PLC.Axis[1].OperationStart,
	Distance := PLC.Axis[1].OperationDistance,
	Velocity := PLC.Axis[1].OperationSpeed,
	Acceleration := PLC.Axis[1].Acceleration,
	Deceleration := PLC.Axis[1].Deceleration,
	Done => PLC.Axis[1].OperationDone);

FB_Relative[2]( //Eixo 2
	Axis := Axis2,
	Execute := PLC.Axis[2].OperationStart,
	Distance := PLC.Axis[2].OperationDistance,
	Velocity := PLC.Axis[2].OperationSpeed,
	Acceleration := PLC.Axis[2].Acceleration,
	Deceleration := PLC.Axis[2].Deceleration,
	Done => PLC.Axis[2].OperationDone);

FB_Relative[3]( //Eixo 1
	Axis := Axis3,
	Execute := PLC.Axis[3].OperationStart,
	Distance := PLC.Axis[3].OperationDistance,
	Velocity := PLC.Axis[3].OperationSpeed,
	Acceleration := PLC.Axis[3].Acceleration,
	Deceleration := PLC.Axis[3].Deceleration,
	Done => PLC.Axis[3].OperationDone);

                    
END_ACTION

ACTION Circular:
                      FB_Circular(
	Axis0 := Axis1,
	Axis1 := Axis2,
	Exec := PLC.OperationCirleStart,
	Circle_Mode := 0,
	CircleRadiual := 0,
	AuxPos := PLC.OperationAuxPos,
	EndPos := PLC.OperationEndPos,
	CircleRadiual := 0,
	Velocity := PLC.Axis[1].OperationSpeed,
	Acceleration := PLC.Axis[1].Acceleration,
	Deceleration := PLC.Axis[1].Deceleration,
	Done => PLC.OperationCircleDone);
                    
END_ACTION
END_PROGRAM

CONFIGURATION Application
  RESOURCE Application ON PLC
    {attribute 'qualified_only'}
    VAR_GLOBAL  (* PLC *)
      Machine : States;  (* Estado da maquina *)
      Safety_Enabled : BOOL;  (* Maquina habilitada *)
      Alarm_Machine : INT;  (* Alarme na máquina *)
      Axis : ARRAY[1..4] OF AxisStruct;  (* Estrutura dos eixos *)
      FB_Homing : ARRAY[1..4] OF SMC_Homing;  (* Bloco de função Homing *)
      IO : IO;  (* Estrutura das entradas digitais *)
      RectangularPieces : ARRAY[0..19] OF Creation_RectanglePoints;  (* Array das posições das peças retangulares *)
      OrthogonalPieces : ARRAY[0..41] OF Creation_OrthogonalPoints;  (* Array das posições das peças ortogonais *)
      CornerPieces : ARRAY[0..8] OF Creation_CornerPoints;  (* Array de posições das peças em L *)
      CornerSquares : ARRAY[0..3] OF Creation_RectanglePoints;
      FormsSquare : Creation_RectanglePoints;  (* Posições das peças retangulares *)
      FormsCircle : Creation_CirclePoints;  (* Posições das peças circulares *)
      FormsHexagon : Creation_HexagonPoints;  (* Posições das peças hexagonais *)
      FormsTriangle : Creation_TranglePoints;  (* Posições das peças triangulares *)
      CutPiece : INT;  (* Peça sendo cortada *)
      CutLine : INT;  (* Linha sendo cortada *)
      CutStraight : INT;  (* Reta sendo cortada *)
      GridTable_Step : INT;  (* Passo atual da construção da tabela *)
      CuttingTable90_Step : INT;  (* Passo atual da construção da tabela *)
      CuttingPause : BOOL;  (* Pausa processo de corte *)
      Piece : INT;  (* Peça atual da array; *)
      PieceFigure : INT;  (* Figura atual da array; *)
      Grid : INT;
      GridFigure : INT;
      GridDesigner_Step : INT;
      GridDesigner_LastLine : INT;  (* Ultima linha criada *)
      CornerArea : INT;
      CornerAreaFigure : INT;
      CornerDesigner_LastCornerArea : INT;
      CornerDesigner_Step : INT;
      CreationRectangles_GreatestHeight : REAL;  (* Maior altura entre as peças *)
      CreationRectangles_GreatestWidth : REAL;  (* Maior largura entre as peças *)
      LastPiece : INT;  (* Ultima peça criada *)
      OperationCirleStart : BOOL;  (* Inicia posição circular *)
      OperationCircleDone : BOOL;
      OperationAuxPos : ARRAY[0..1] OF LREAL;
      OperationEndPos : ARRAY[0..1] OF LREAL;
    END_VAR
    {attribute 'qualified_only'}
    VAR_GLOBAL  (* IHM *)
      btStart : BOOL;  (* Botão de start virtual *)
      btStop : BOOL;  (* Botão de stop virtual *)
      btReset : BOOL;  (* Botão de reset virtual *)
      btStartHome : BOOL;  (* Botao de start homing virtual *)
      btGoToZero : BOOL;  (* Botão virtual retorna para ponto zero *)
      btRotateSaw : BOOL;  (* Botão virtual para girar a serra *)
      RotateValue : REAL;  (* Valor para girar a serra *)
      btSetPoint : BOOL;  (* Define novo ponto zero *)
      btTableUp : BOOL;  (* Botão virtual sobe mesa *)
      btTableDown : BOOL;  (* Botão virtual desce mesa *)
      AlarmOn : INT;  (* Alarme na máquina *)
      DeleteLastPiece : BOOL;  (* Deletar ultima peça *)
      FinishPiece : BOOL;  (* Finalizar criação *)
      CancelPiece : BOOL;  (* Cancelar criação *)
      Figure : INT;  (* Figura para seleção *)
      NewWidth : REAL;  (* Largura da nova peça *)
      NewHeight : REAL;  (* Altura da nova peça *)
      ZeroMessage : BOOL;  (* Mensagem de valores zerados na IHM *)
      NoFigure : BOOL;  (* Mensagem de nenhuma figura selecionada *)
      PauseMessage : BOOL;  (* Mensagem de pause na IHM *)
      NoPiece : BOOL;  (* Mensagem nenhuma peça criada *)
      ContinueOperation : BOOL;  (* Continua operação de corte *)
      CutMode : BOOL;  (* Modo de corte *)
      CreationRectangle_Start : BOOL;  (* Iniciar criação de peça retangular *)
      CreationRectangle_MakeNewPieceSide : BOOL;  (* Gerar nova figura em cima *)
      CreationRectangle_MakeNewPieceDown : BOOL;  (* Gerar nova figura em baixo *)
      CreationOrthogonal_MakeOrthogonal : BOOL;  (* Gerar nova figura ortogonal *)
      CreationOrthogonal_Start : BOOL;  (* Iniciar criação de peça ortogonal *)
      CreationOrthogonal_GridLines : INT;  (* Quantidade de linhas do corte ortogonal *)
      CreationOrthogonal_GridColumns : INT;  (* Quantidade de colunas do corte ortogonal *)
      CreationCorner_Start : BOOL;  (* Inicia criação de peça em L *)
      CreationCorner_MakeCorner : BOOL;  (* Gerar nova figura em L *)
      CreationCorner_X1 : REAL;  (* Tamanho X1 da peça L *)
      CreationCorner_X2 : REAL;  (* Tamanho X2 da peça L *)
      CreationCorner_Y1 : REAL;  (* Tamanho Y1 da peça L *)
      CreationCorner_Y2 : REAL;  (* Tamanho Y2 da peça L *)
      CreationCorner_ReverseCorner : BOOL;  (* Inverter corte L *)
      CreationCorner_CornerDisplacement : REAL;  (* Distancia entre peças L *)
      CreationCorner_MirrorCorner : BOOL;  (* Espelhamento de corte L *)
      CreationForms_Start : BOOL;  (* Inicia criação de peça em formas *)
      CreationForms_MakeNewPiece : BOOL;  (* Gerar nova figura *)
      CreationForms_Width : REAL;  (* Posição do centro do circulo em X *)
      CreationForms_Height : REAL;  (* Posição do centro do circulo em Y *)
      CreationForms_Radius : REAL;  (* Raio do circulo *)
      CreationForms_Perimeter : REAL;  (* Perimetro do hexagono *)
      Axis : ARRAY[1..4] OF AxisStruct;
      Input : ARRAY[0..15] OF BOOL;
      PrZeroPieceMachineX : REAL;  (* Zero peça em X *)
      PrZeroPieceMachineY : REAL;  (* Zero peça em Y *)
      PrEntryEdgeX : REAL;  (* Borda de entrada *)
      PrEntryEdgeY : REAL;  (* Borda de entrada *)
      PrReverseCornerEntryX : REAL;  (* Borda interna L invertido *)
      PrReverseCornerEntryY : REAL;  (* Borda interna L invertido *)
      PrCornerEdgeX : REAL := 95;  (* Borda interna *)
      PrCornerEdgeY : REAL := 90;  (* Borda interna *)
      PrLeadingEdgeX : REAL;  (* Borda de saida *)
      PrLeadingEdgeY : REAL;  (* Borda de saida *)
      PrOutsidePiece : REAL;  (* Posição fora da peça *)
      PrInsidePiece : REAL;  (* Posição dentro da peça *)
      SawThickness : REAL := 3.4;  (* Espessura da serra *)
    END_VAR
    TASK MainTask(INTERVAL := T#2ms, PRIORITY := 0);
    TASK MotionTask(INTERVAL := T#0.5ms, PRIORITY := 1);
    TASK EtherCAT_Task(INTERVAL := T#0.5ms, PRIORITY := 1);
    PROGRAM Main WITH MainTask : Main;
    PROGRAM POU WITH MainTask : POU;
    PROGRAM Motion WITH MotionTask : Motion;
  END_RESOURCE
END_CONFIGURATION
